Fanuc KAREL source: ks00018.KL

-- PROVISIONAL review KL for V1013-1; original PC SHA256 7d790a00119560c65ad49774b4dc748296aae7ebdac467764dc9f26bec6f13c2
-- Incomplete behavior may be omitted. Consult companion uncertainty JSON. Do not deploy.
PROGRAM KS00018
%NOLOCKGROUP
VAR
  A : FILE
  B : FILE
  FLAG : BOOLEAN
  N : INTEGER
  STATUS : INTEGER
  PN : STRING[80]
  VN : STRING[80]
BEGIN
  -- UNRESOLVED_PC offsets 5-13; opcodes 3F,75
  -- UNRESOLVED_PC offsets 18-27; opcodes 3F,75
  -- UNRESOLVED_PC offsets 32-47; opcodes 22,63,23
  -- UNRESOLVED_PC offsets 52-56; opcodes 7F
END KS00018
